(* IEC 61131-3 sources: rusty/tests/lit/single/types, 3 files *)

(* ---- self_referential_pointer_to.st ---- *)
// RUN: %COMPILE %s && %RUN | %CHECK %s

// Test self-referential struct broken by POINTER TO
TYPE LinkedList : STRUCT
    value : DINT;
    next : POINTER TO LinkedList;
END_STRUCT END_TYPE

FUNCTION main : DINT
    VAR
        list1 : LinkedList;
        list2 : LinkedList;
    END_VAR

    list1.value := 10;
    list2.value := 20;

    // Link them together
    list1.next := ADR(list2);
    list2.next := ADR(list1);

    // CHECK: List1 value: 10
    printf('List1 value: %d$N', list1.value);

    // CHECK: List2 value: 20
    printf('List2 value: %d$N', list2.value);

    main := 0;
END_FUNCTION

(* ---- self_referential_ref_to.st ---- *)
// RUN: %COMPILE %s && %RUN | %CHECK %s

// Test self-referential struct broken by REF_TO
TYPE TreeNode : STRUCT
    data : DINT;
    left : REF_TO TreeNode;
    right : REF_TO TreeNode;
END_STRUCT END_TYPE

FUNCTION main : DINT
    VAR
        root : TreeNode;
        leftChild : TreeNode;
        rightChild : TreeNode;
    END_VAR

    root.data := 50;
    leftChild.data := 25;
    rightChild.data := 75;

    // Build tree structure
    root.left := REF(leftChild);
    root.right := REF(rightChild);

    // CHECK: Root: 50
    printf('Root: %d$N', root.data);

    // CHECK: Left: 25
    printf('Left: %d$N', root.left^.data);

    // CHECK: Right: 75
    printf('Right: %d$N', root.right^.data);

    main := 0;
END_FUNCTION

(* ---- self_referential_struct_via_reference.st ---- *)
// RUN: %COMPILE %s && %RUN | %CHECK %s

TYPE Node : STRUCT
    data : DINT;
    next : REFERENCE TO Node;
END_STRUCT END_TYPE

FUNCTION main : DINT
    VAR
        node1 : Node;
        node2 : Node;
    END_VAR

    node1.data := 42;
    node2.data := 84;

    // Create circular reference
    node1.next REF= node2;
    node2.next REF= node1;

    // CHECK: Node1 data: 42
    printf('Node1 data: %d$N', node1.data);

    // CHECK: Node2 data: 84
    printf('Node2 data: %d$N', node2.data);

    // CHECK: Node1->next->data: 84
    printf('Node1->next->data: %d$N', node1.next.data);

    // CHECK: Node2->next->data: 42
    printf('Node2->next->data: %d$N', node2.next.data);

    // CHECK: Circular reference works: 42
    printf('Circular reference works: %d$N', node1.next.next.data);

    main := 0;
END_FUNCTION
